// TwinCAT 3 PLC project TcToolkitSample2_PLC
// ProgramVersion: 3.1.4024.0
// libraries:
//   Tc2_Standard, * (Beckhoff Automation GmbH)
//   Tc2_System, * (Beckhoff Automation GmbH)
//   Tc3_Module, * (Beckhoff Automation GmbH)
// project tree:
//   GVLs/ GVL_Main.TcGVL
//   / PlcTask.TcTTO
//   POUs/ MAIN.TcPOU, FB_Valve.TcPOU, FB_Cylinder.TcPOU
//   DUTs/ E_ValveState.TcDUT, ST_TankData.TcDUT
//   POUs/Interfaces/ I_Valve.TcIO

CONFIGURATION TcToolkitSample2_PLC
    RESOURCE PLC ON TwinCAT3
        TASK PlcTask(INTERVAL := T#10ms, PRIORITY := 20);
        PROGRAM MAIN WITH PlcTask : MAIN;
    END_RESOURCE
END_CONFIGURATION

// ---- DUTs/E_ValveState.TcDUT
TYPE E_ValveState :
(
	Closed := 0,
	Opening := 1,
	Open := 2,
	Closing := 3
);
END_TYPE

// ---- DUTs/ST_TankData.TcDUT
TYPE ST_TankData :
STRUCT
	fLevel		: LREAL;
	fSetpoint	: LREAL := 50.0;
	eInlet		: E_ValveState;
	bAlarm		: BOOL;
END_STRUCT
END_TYPE

// ---- GVLs/GVL_Main.TcGVL
{attribute 'qualified_only'}
VAR_GLOBAL
	stTank		: ST_TankData;
	nCycles		: UDINT;
	bFillRequest	: BOOL;
END_VAR

// ---- POUs/Interfaces/I_Valve.TcIO
INTERFACE I_Valve

METHOD Open : BOOL
END_METHOD

PROPERTY State : E_ValveState
GET
END_GET
SET
END_SET
END_PROPERTY

END_INTERFACE

// ---- POUs/MAIN.TcPOU
PROGRAM MAIN
VAR
	fbValve		: FB_Valve;
	ipValve		: I_Valve;
	fbCylinder	: FB_Cylinder;
	nStroke		: UINT;
END_VAR

GVL_Main.nCycles := GVL_Main.nCycles + 1;
ipValve := fbValve;
IF GVL_Main.bFillRequest AND GVL_Main.stTank.fLevel < GVL_Main.stTank.fSetpoint THEN
	ipValve.Open();
END_IF
fbValve(bClose := GVL_Main.stTank.fLevel >= GVL_Main.stTank.fSetpoint);
GVL_Main.stTank.eInlet := fbValve.State;
GVL_Main.stTank.bAlarm := GVL_Main.stTank.eInlet = E_ValveState.Open AND NOT fbValve.bIsOpen;
fbCylinder(bExtend := fbValve.bIsOpen);
nStroke := fbCylinder.Stroke();

END_PROGRAM

// ---- POUs/FB_Valve.TcPOU
FUNCTION_BLOCK FB_Valve IMPLEMENTS I_Valve
VAR_INPUT
	bClose	: BOOL;
END_VAR
VAR_OUTPUT
	bIsOpen	: BOOL;
END_VAR
VAR
	_eState	: E_ValveState;
	_nTicks	: UINT;
END_VAR

IF bClose THEN
	Act_Close();
END_IF
IF _eState = E_ValveState.Opening THEN
	_nTicks := _nTicks + 1;
	IF _nTicks >= 10 THEN
		_eState := E_ValveState.Open;
	END_IF
END_IF
bIsOpen := _eState = E_ValveState.Open;

METHOD Open : BOOL
VAR
END_VAR
IF _eState = E_ValveState.Closed THEN
	_eState := E_ValveState.Opening;
	_nTicks := 0;
END_IF
Open := _eState <> E_ValveState.Closed;
END_METHOD

PROPERTY State : E_ValveState
GET
State := _eState;
END_GET
SET
_eState := State;
END_SET
END_PROPERTY

ACTION Act_Close:
_eState := E_ValveState.Closed;
_nTicks := 0;
END_ACTION

END_FUNCTION_BLOCK

// ---- POUs/FB_Cylinder.TcPOU
FUNCTION_BLOCK FB_Cylinder
VAR_INPUT
	bExtend		: BOOL;
	nStrokeTicks	: UINT := 5;
END_VAR
VAR_OUTPUT
	bExtended	: BOOL;
END_VAR
VAR
	_nTicks	: UINT;
END_VAR

IF bExtend THEN
	IF _nTicks < nStrokeTicks THEN
		_nTicks := _nTicks + 1;
	END_IF
ELSE
	_nTicks := 0;
END_IF
bExtended := bExtend AND _nTicks >= nStrokeTicks;

METHOD Stroke : UINT
VAR
END_VAR
Stroke := _nTicks;
END_METHOD

END_FUNCTION_BLOCK
